Fanuc KAREL source: kb00187.KL

-- PROVISIONAL review KL for V770-1; original PC SHA256 384dc920c64fc260a660a8db7b2891b88a136894a2ec7a510ce11c4b31a756a8
-- Incomplete behavior may be omitted. Consult companion uncertainty JSON. Do not deploy.
PROGRAM KB00187
%NOLOCKGROUP
VAR
  P1 : REAL
  RESULT : REAL
BEGIN
  -- UNRESOLVED_PC offsets 5-16; opcodes 2E,23
  -- UNRESOLVED_PC offsets 21-36; opcodes 27,22,76,23
  -- UNRESOLVED_PC offsets 41-45; opcodes 7F
END KB00187
